TYPE "ST_PressDemoParCmd"
VERSION : 0.1
   STRUCT
      "Reserved" : Bool;
   END_STRUCT;
END_TYPE
